INTERFACE I_Motor

METHOD Update
VAR_INPUT
    run : BOOL;
    delay : TIME;
END_VAR
END_METHOD

PROPERTY SpeedSetpoint : LREAL
GET
END_GET
SET
END_SET
END_PROPERTY

PROPERTY Running : BOOL
GET
END_GET
END_PROPERTY

PROPERTY Faulted : BOOL
GET
END_GET
END_PROPERTY

PROPERTY ActualSpeed : LREAL
GET
END_GET
END_PROPERTY

END_INTERFACE

(* stored: Version 1.1.0.1, ProductVersion 3.1 *)
